// TIA Portal project "tanque_sensor_temperatura_V2" (V12)

(* hardware
DEVICE "S7-1200 station_1"  SIMATIC 1200-Station
   slot 0: "S7-1200 rack"  Rack  V1.0
   slot 1: "PLC_1"  CPU 1214C DC/DC/DC  6ES7 214-1AG31-0XB0  V3.0
DEVICE "HMI_1"  KTP600 Basic color PN
   slot 0: "HMI"  HMI  6AV6647-0AD11-3AX0  12.0.0.0
   slot 1: "HMI_RT_1"  KTP600 Basic color PN  6AV6647-0AD11-3AX0  12.0.0.0
   slot 5: "HMI_1.IE_CP_1"  PROFINET Interface
      slot 1: "PROFINET Interface_1"  PROFINET Interface
         slot 1: "Port_1"  Port
DEVICE "S7-1200 station_2"  SIMATIC 1200-Station
   slot 0: "S7-1200 rack"  Rack  V1.0
   slot 1: "PLC_2"  CPU 1214C DC/DC/DC  6ES7 214-1AG31-0XB0  V3.0
DEVICE "HMI_2"  KTP600 Basic color PN
   slot 0: "HMI"  HMI  6AV6647-0AD11-3AX0  12.0.0.0
   slot 1: "HMI_RT_2"  KTP600 Basic color PN  6AV6647-0AD11-3AX0  12.0.0.0
   slot 5: "HMI_2.IE_CP_1"  PROFINET Interface
      slot 1: "PROFINET Interface_1"  PROFINET Interface
         slot 1: "Port_1"  Port
*)

// ===== PLC "PLC_1"  CPU 1214C DC/DC/DC =====

VAR_GLOBAL   // PLC tag table "Default tag table"
   "resistor" AT %Q0.2 : Bool;
   "sensor temp" AT %Q0.3 : Bool;
END_VAR

VAR_GLOBAL   // PLC tag table "Tag table_1"
   "liga" AT %I0.0 : Bool;
   "desliga" AT %I0.1 : Bool;
   "s1" AT %I0.2 : Bool;   // s1 T Nvb
   "s2" AT %I0.3 : Bool;   // s2 T Nva
   "s3" AT %I0.4 : Bool;   // s3 Ts Nvb
   "s4" AT %I0.5 : Bool;   // s4 Ts Nva
   "motor" AT %Q0.0 : Bool;
   "solenoide" AT %Q0.1 : Bool;
   "sistema" AT %M0.0 : Bool;
   "emergencia" AT %I0.6 : Bool;
   "valor sensor tensão" AT %IW64 : Int;
   "valor sensor digital" AT %MD0 : Real;
   "valor sensor graus" AT %MW4 : UInt;
   "liga resistor" AT %I0.7 : Bool;
   "prioridade solenoide" AT %M0.1 : Bool;
   "temperatura IHM" AT %MD2 : UDInt;
   "selo resistor" AT %M0.2 : Bool;
   "fluxo motor" AT %M0.3 : Bool;
   "fluxo solenoide" AT %M6.0 : Bool;
END_VAR

// folder: System blocks/Program resources

DATA_BLOCK "IEC_Timer_0_DB_1"   // DB2
{ S7_Optimized_Access := 'FALSE' }
AUTHOR : Simatic
FAMILY : IEC
NAME : IEC_TMR
VERSION : 1.0
// stored: InstanceOfName ?
"?"
BEGIN
END_DATA_BLOCK

// folder: (top level)

ORGANIZATION_BLOCK "Main"   // OB1, LAD, ProgramCycle
TITLE = "Main Program Sweep (Cycle)"
{ S7_Optimized_Access := 'FALSE' }
VERSION : 0.1
   VAR_TEMP   // added for the SCL form of the ladder/FBD networks
      _w1 : Bool;
   END_VAR
BEGIN

REGION Network 1
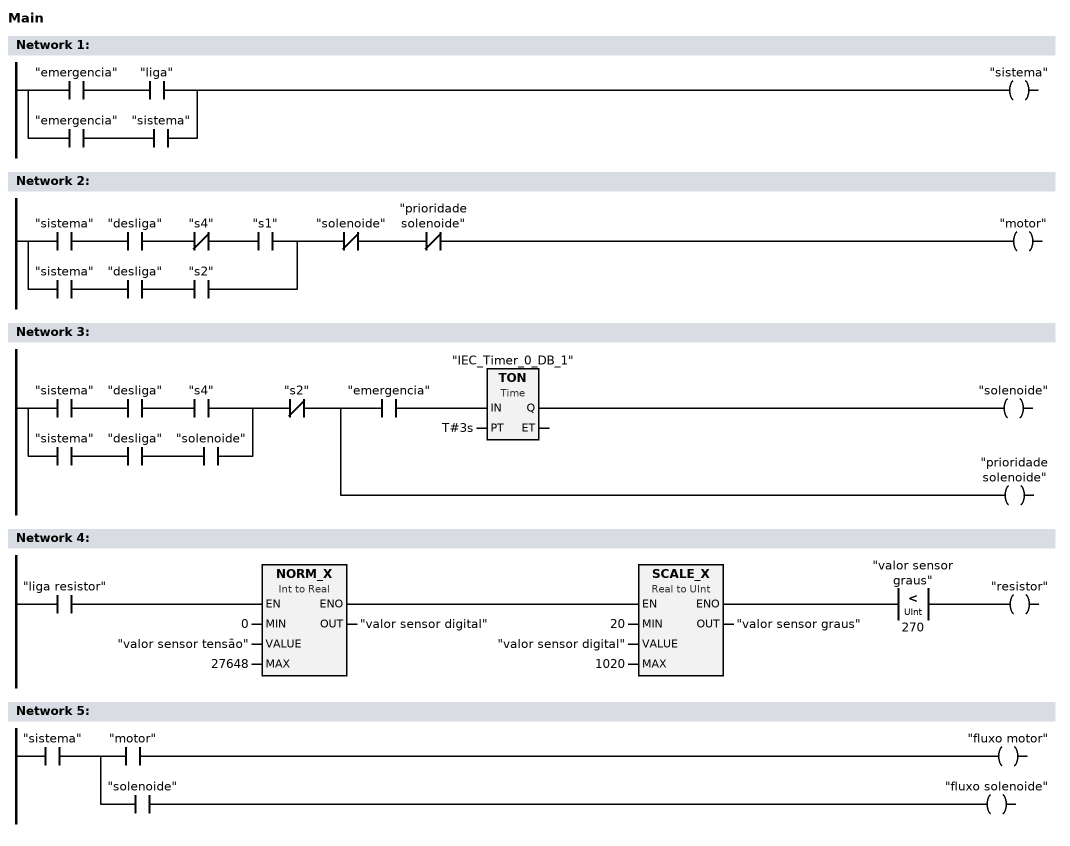
   RUNG wire#powerrail
      Contact( "emergencia" )
      Contact( "liga" )
      wire#w1
      Coil( "sistema" )
   END_RUNG
   RUNG wire#powerrail
      Contact( "emergencia" )
      Contact( "sistema" )
   END_RUNG wire#w1
   // the same network as SCL:
   "sistema" := ("emergencia" AND "liga") OR ("emergencia" AND "sistema");
END_REGION

REGION Network 2
   RUNG wire#powerrail
      Contact( "sistema" )
      Contact( "desliga" )
      I_Contact( "s4" )
      Contact( "s1" )
      wire#w1
      I_Contact( "solenoide" )
      I_Contact( "prioridade solenoide" )
      Coil( "motor" )
   END_RUNG
   RUNG wire#powerrail
      Contact( "sistema" )
      Contact( "desliga" )
      Contact( "s2" )
   END_RUNG wire#w1
   // the same network as SCL:
   "motor" := (("sistema" AND "desliga" AND NOT "s4" AND "s1") OR ("sistema" AND "desliga" AND "s2")) AND NOT "solenoide" AND NOT "prioridade solenoide";
END_REGION

REGION Network 3
   #_w1 := (("sistema" AND "desliga" AND "s4") OR ("sistema" AND "desliga" AND "solenoide")) AND NOT "s2";
   "IEC_Timer_0_DB_1".TON(IN := #_w1 AND "emergencia", PT := T#3s);
   "solenoide" := "IEC_Timer_0_DB_1".Q;
   "prioridade solenoide" := #_w1;
END_REGION

REGION Network 4
   RUNG wire#powerrail
      Contact( "liga resistor" )
      { S7_Templates := "[SrcType := Int, DestType := Real]"; S7_GenerateENO := "TRUE" } Normalize(min := 0, value := "valor sensor tensão", max := 27648, out => "valor sensor digital")
      { S7_Templates := "[SrcType := Real, DestType := UInt]"; S7_GenerateENO := "TRUE" } Scale(min := 20, value := "valor sensor digital", max := 1020, out => "valor sensor graus")
      { S7_Templates := "SrcType := UInt" } LT_Contact(in1 := "valor sensor graus", in2 := 270)
      Coil( "resistor" )
   END_RUNG
   // the same network as SCL:
   // ENO of a box is taken as its EN; it also drops when the box reports an error
   IF "liga resistor" THEN
       "valor sensor digital" := NORM_X(MIN := 0, VALUE := "valor sensor tensão", MAX := 27648);
       "valor sensor graus" := SCALE_X(MIN := 20, VALUE := "valor sensor digital", MAX := 1020);
   END_IF;
   "resistor" := "liga resistor" AND ("valor sensor graus" < 270);
END_REGION

REGION Network 5
   RUNG wire#powerrail
      Contact( "sistema" )
      wire#w1
      Contact( "motor" )
      Coil( "fluxo motor" )
   END_RUNG
   RUNG wire#w1
      Contact( "solenoide" )
      Coil( "fluxo solenoide" )
   END_RUNG
   // the same network as SCL:
   "fluxo motor" := "sistema" AND "motor";
   "fluxo solenoide" := "sistema" AND "solenoide";
END_REGION
END_ORGANIZATION_BLOCK

// ===== PLC "PLC_2"  CPU 1214C DC/DC/DC =====

VAR_GLOBAL   // PLC tag table "Default tag table"
   "RT" AT %I0.0 : Bool;
   "B0" AT %I0.1 : Bool;
   "B1" AT %I0.2 : Bool;
   "M1" AT %Q0.0 : Bool;
END_VAR

ORGANIZATION_BLOCK "Main"   // OB1, LAD, ProgramCycle
TITLE = "Main Program Sweep (Cycle)"
{ S7_Optimized_Access := 'FALSE' }
VERSION : 0.1
BEGIN

REGION Network 1: Liga Desliga
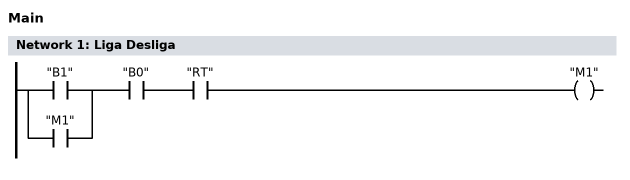
   RUNG wire#powerrail
      Contact( "B1" )
      wire#w1
      Contact( "B0" )
      Contact( "RT" )
      Coil( "M1" )
   END_RUNG
   RUNG wire#powerrail
      Contact( "M1" )
   END_RUNG wire#w1
   // the same network as SCL:
   "M1" := ("B1" OR "M1") AND "B0" AND "RT";
END_REGION
END_ORGANIZATION_BLOCK

(* ===== HMI "HMI_RT_1" =====
connection "HMI_connection_1": ETHERNET, SMART_S7_1200_OMS

HMI tags "Tag table_1"
   "s1" : Bool = PLC "s1", 100 ms
   "s2" : Bool = PLC "s2", 100 ms
   "s3" : Bool = PLC "s3", 100 ms
   "s4" : Bool = PLC "s4", 100 ms
   "HMI_desliga" : Bool = PLC "sistema", 100 ms
   "HMI_liga" : Bool = PLC "sistema", 100 ms
   "solenoide" : Bool = PLC "solenoide", 100 ms
   "motor" : Bool = PLC "motor", 100 ms
   "solenoide_1" : Bool, 1 s

screen "TELA INICIAL" 320x240, template "Template_1"
   TextField "HmiScreenItemData_2" at 20,0 size 256x17

screen "SISTEMA" 320x240, template "Template_1"
   TextField "HmiScreenItemData" at 32,-1 size 256x17

screen "DOCUMENTAÇÃO" 320x240, template "Template_1"
   TextField "HmiScreenItemData" at 27,0 size 256x17
   GraphicView "Graphic view_1" at 0,0 size 320x206
   Button "Button_1" at 13,199 size 137x37
   Button "Button_2" at 186,203 size 128x32

screen "Different jobs" 320x240, template "Template_1"
   Button "HmiScreenItemData" at 1,32 size 104x30
   Button "HmiScreenItemData_1" at 1,63 size 104x30
   Button "HmiScreenItemData_2" at 1,94 size 104x30
   Button "HmiScreenItemData_3" at 1,125 size 104x30
   Button "HmiScreenItemData_4" at 1,156 size 104x30
   Button "HmiScreenItemData_5" at 1,1 size 104x30
*)

(* ===== HMI "HMI_RT_2" =====
connection "HMI_connection_2": ETHERNET, SMART_S7_1200_OMS

screen "TELA INICIAL" 320x240, template "Template_1"
   TextField "HmiScreenItemData_2" at 35,6 size 256x17

screen "DOCUMENTAÇÃO" 320x240, template "Template_1"
   TextField "HmiScreenItemData" at 34,3 size 256x17

screen "SISTEMAS" 320x240, template "Template_1"
   TextField "HmiScreenItemData" at 36,3 size 256x17
*)